(* IEC 61131-3 sources: plc-sbom-builder/samples/maschine-xy/programm/Roboterzelle/POUs, 1 file *)

(* ---- MAIN.st ---- *)
PROGRAM MAIN
VAR
    fTemperatur : LREAL;
END_VAR

fTemperatur := 21.5;
